// TIA Portal V21 export
// export: Created 2026-10-08T12:30:16.9154675Z, ExportSetting WithDefaults, DisplayName Totally Integrated Automation Portal, DisplayVersion V21 Update 2, DisplayName TIA Portal Test Suite Advanced, DisplayVersion V21, DisplayName SINAMICS Startdrive Advanced, DisplayVersion V21 HF2, DisplayName SINAMICS DCC, DisplayVersion V21, DisplayName SINAMICS Startdrive G110M, G120, G120C, G120D, G120P, G115D, DisplayVersion V21 HF2, DisplayName SINAMICS Startdrive G130, G150, S120, S150, G200, G220, S200, S210, S220, Innomotics MVD, DisplayVersion V21 HF2, DisplayName STEP 7 Professional, DisplayVersion V21 Update 2, DisplayName STEP 7 Safety, DisplayVersion V21, DisplayName Tech WebApplication, DisplayVersion V21, DisplayName WinCC Basic/Comfort/Advanced, DisplayVersion V21 Update 2, DisplayName WinCC Unified, DisplayVersion V21 Update 2
FUNCTION_BLOCK "Tgp_NumericFB_LAD"   // FB57, LAD
{ S7_Optimized_Access := 'TRUE' }
VERSION : 0.1
// stored: AutoNumber true, IsIECCheckEnabled false, IsRetainMemResEnabled false, MemoryReserve 100, SetENOAutomatically false, UDAEnableTagReadback false
   VAR_INPUT
      Enable : Bool;
      Delta : Int;
      Reset : Bool;
   END_VAR
   VAR_OUTPUT
      Total : Int;
   END_VAR
   VAR_IN_OUT
      Accumulator : Int;
   END_VAR
   VAR
      Child { S7_SetPoint := 'True'} : "Tgp_NumericFB";
   END_VAR
BEGIN

REGION Network 1
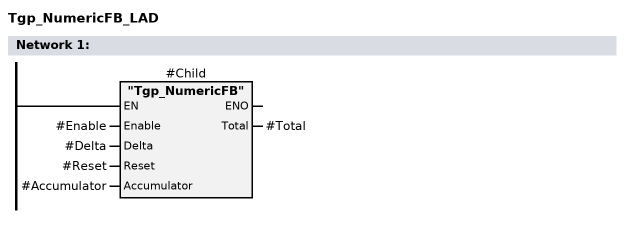
   RUNG wire#powerrail
      #Child(Enable := #Enable, Delta := #Delta, Reset := #Reset, Accumulator := #Accumulator, Total => #Total)
   END_RUNG
   // the same network as SCL:
   #Child(Enable := #Enable, Delta := #Delta, Reset := #Reset, Accumulator := #Accumulator, Total => #Total);   // "Tgp_NumericFB"
END_REGION
END_FUNCTION_BLOCK
